SUBAPPLICATION Uebung_OPC_L18_AX (* Objekte/Variablen per PUBLISH_0: I1 CREATE_OBJECT, I2 CREATE_VARIABLE, I3 DELETE_VARIABLE, I4 DELETE_OBJECT - lokal auf einem Geraet *)
  (* Standard: 61499-2; Description: Copyright (c) 2026 Meisterschulen am Ostbahnhof This program and the accompanying materials are made available under the terms of the Eclipse Public License 2.0 which is available at https://www.eclipse.org/legal/epl-2.0/ SPDX-License-Identifier: EPL-2.0 *)
  (* Version 1.0, 2026-10-18, Franz Höpfinger, Meisterschulen am Ostbahnhof, opcua.adoc-Beispiel lokal (Meins/OPC_UA_Lokal) *)
  PACKAGE Meins::OPC_UA_Lokal;
  IMPORT Meins::OPC_UA_Lokal::const::OpcUaLokal::L18_OBJ_CREATE;
  IMPORT Meins::OPC_UA_Lokal::const::OpcUaLokal::L18_VAR_CREATE;
  IMPORT Meins::OPC_UA_Lokal::const::OpcUaLokal::L18_VAR_DELETE;
  IMPORT Meins::OPC_UA_Lokal::const::OpcUaLokal::L18_OBJ_DELETE;
  IMPORT logiBUS::io::DI::logiBUS_DI::Input_I1;
  IMPORT logiBUS::io::DI::logiBUS_DI::Input_I2;
  IMPORT logiBUS::io::DI::logiBUS_DI::Input_I3;
  IMPORT logiBUS::io::DI::logiBUS_DI::Input_I4;
  IMPORT logiBUS::io::DI::logiBUS_DI_Events::BUTTON_PRESS_DOWN;
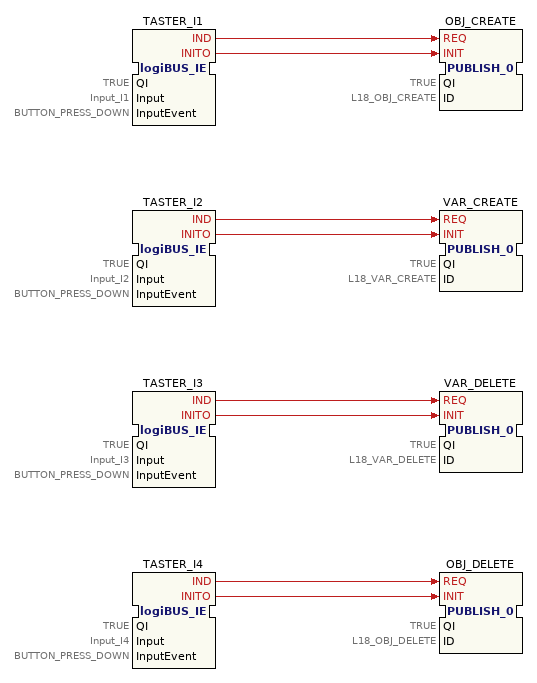
  FBS
    TASTER_I1 : logiBUS::io::DI::logiBUS_IE(QI := TRUE, Input := Input_I1, InputEvent := BUTTON_PRESS_DOWN);
    OBJ_CREATE : iec61499::net::PUBLISH_0(QI := TRUE, ID := L18_OBJ_CREATE);
    TASTER_I2 : logiBUS::io::DI::logiBUS_IE(QI := TRUE, Input := Input_I2, InputEvent := BUTTON_PRESS_DOWN);
    VAR_CREATE : iec61499::net::PUBLISH_0(QI := TRUE, ID := L18_VAR_CREATE);
    TASTER_I3 : logiBUS::io::DI::logiBUS_IE(QI := TRUE, Input := Input_I3, InputEvent := BUTTON_PRESS_DOWN);
    VAR_DELETE : iec61499::net::PUBLISH_0(QI := TRUE, ID := L18_VAR_DELETE);
    TASTER_I4 : logiBUS::io::DI::logiBUS_IE(QI := TRUE, Input := Input_I4, InputEvent := BUTTON_PRESS_DOWN);
    OBJ_DELETE : iec61499::net::PUBLISH_0(QI := TRUE, ID := L18_OBJ_DELETE);
  END_FBS
  EVENT_CONNECTIONS
    TASTER_I1.IND TO OBJ_CREATE.REQ;
    TASTER_I1.INITO TO OBJ_CREATE.INIT;
    TASTER_I2.IND TO VAR_CREATE.REQ;
    TASTER_I2.INITO TO VAR_CREATE.INIT;
    TASTER_I3.IND TO VAR_DELETE.REQ;
    TASTER_I3.INITO TO VAR_DELETE.INIT;
    TASTER_I4.IND TO OBJ_DELETE.REQ;
    TASTER_I4.INITO TO OBJ_DELETE.INIT;
  END_CONNECTIONS
END_SUBAPPLICATION
